TYPE U_DWORD_REAL1 :
UNION
	dw : DWORD;
    out  : REAL;
END_UNION
END_TYPE

(* stored: Version 1.1.0.1
   DUT U_DWORD_REAL1: Id {0f3c4c2d-2ec1-498c-88a7-cfab8749de75} *)
